(* CODESYS project Signals.xml

Project tree, tasks and I/O mapping:
  program Signals [LD]
*)

// Signals
PROGRAM Signals
VAR
	TON_0: TON;
	TON_1: TON;
	tSignalTime:TIME:=T#1S;
	BLINK_0: BLINK;
END_VAR

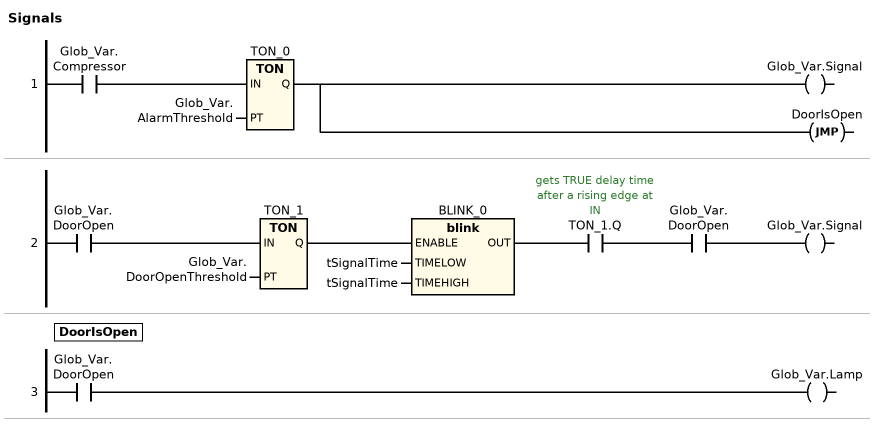
// NETWORK 1
TON_0(IN := Glob_Var.Compressor, PT := Glob_Var.AlarmThreshold); // TON
Glob_Var.Signal := TON_0.Q;
IF TON_0.Q THEN JMP DoorIsOpen; END_IF

// NETWORK 2
//   TON_1.Q: gets TRUE delay time after a rising edge at IN
TON_1(IN := Glob_Var.DoorOpen, PT := Glob_Var.DoorOpenThreshold); // TON
BLINK_0(ENABLE := TON_1.Q, TIMELOW := tSignalTime, TIMEHIGH := tSignalTime); // blink
Glob_Var.Signal := BLINK_0.OUT AND TON_1.Q AND Glob_Var.DoorOpen;

// NETWORK 3
DoorIsOpen:
Glob_Var.Lamp := Glob_Var.DoorOpen;

END_PROGRAM
